Fanuc KAREL source: kb00197.KL

-- PROVISIONAL review KL for V940-1; original PC SHA256 4230892b2e8468a453491833a6e3494f1c4426453fac8a098819c032b0ee426d
-- Incomplete behavior may be omitted. Consult companion uncertainty JSON. Do not deploy.
PROGRAM KB00197
%NOLOCKGROUP
BEGIN
  -- V9_ZERO_TABLE_METADATA_HINT layout=0002_ascii; no indexed target words; source/name/runtime held
  -- UNRESOLVED_PC offsets 5-14; opcodes 3F,75
  -- UNRESOLVED_PC offsets 19-26; opcodes 9D,23
  -- UNRESOLVED_PC offsets 31-38; opcodes 9D,23
  -- UNRESOLVED_PC offsets 43-73; opcodes 27,22,22,2A,22,22,31
  -- UNRESOLVED_PC offsets 78-82; opcodes 7F
END KB00197
